(* PLC project probe.project, CODESYS CODESYS V3.5 SP17 Patch 3 *)
(* stored: creationDateTime 2026-10-20T03:54:26.8891721, modificationDateTime 1601-01-01T03:00:00 *)

PROGRAM PRG_ProbeMain
  VAR
    fbSt : FB_ProbeSt;
    fbFbd : FB_ProbeFbd;
    fbLd : FB_ProbeLd;
    fbFbdEno : FB_ProbeFbdEno;
    fbCfc : FB_ProbeCfc;
    fbPcfc : FB_ProbePcfc;
    fbOop : FB_ProbeOop2;
    fbIl : FB_ProbeIl;
    stVal : ST_ProbeVal;
  END_VAR

            fbSt(xIn := GVL_ProbeP.xFlag);
fbFbd(rLevel := 1.0, rHigh := 0.5, xEnable := TRUE);
fbLd(xStart := GVL_ProbeP.xFlag);
fbFbdEno(xEn := TRUE, iSp := 5);
fbCfc(rIn := 1.0, rLo := 0.0, rHi := 10.0);
fbPcfc(rA := 2.0, rK := 3.0);
fbOop(xIn := TRUE);
fbIl(xIn := TRUE, iN := 3);
GVL_ProbeP.diHours := GVL_ProbeP.diHours + 1;
stVal.eMode := E_ProbeMode.Auto;

          
END_PROGRAM
